// TIA Portal V20 export
// export: Created 2026-10-24T18:20:57.3148607Z, ExportSetting WithDefaults, DisplayName Totally Integrated Automation Portal, DisplayVersion V20 Update 6, DisplayName TIA Portal Openness, DisplayVersion V20 Update 6, DisplayName TIA Portal Version Control Interface, DisplayVersion V20 Update 6, DisplayName SINAMICS Startdrive Advanced, DisplayVersion V20 SP1 Update 2, DisplayName SINAMICS Startdrive G110M, G120, G120C, G120D, G120P, G115D, DisplayVersion V20 SP1 Update 2, DisplayName SINAMICS Startdrive G130, G150, S120, S150, SINAMICS MV, G220, S200, S210, DisplayVersion V20 SP1 Update 2, DisplayName STEP 7 Professional, DisplayVersion V20 Update 6, DisplayName STEP 7 Safety, DisplayVersion V20 Update 2, DisplayName WinCC Basic/Comfort/Advanced, DisplayVersion V20 Update 6, DisplayName WinCC Unified, DisplayVersion V20 Update 6
TYPE "UDT_Motor"
TITLE = Motor data
// stored: IsFailsafeCompliant false
   STRUCT
      Enable : Bool;   // Release from the line control
      Running : Bool;   // Feedback: motor is running
      Fault : Bool;   // Motor protection tripped
      SpeedSetpoint : Real := 1450.0;   // Speed setpoint in rpm
      ActualSpeed : Real;   // Measured speed in rpm
      RunTime : Time := T#0MS;   // Accumulated run time
      StartCount : DInt := 0;   // Number of starts
   END_STRUCT;
END_TYPE
